TYPE "ST_PressDemoStationCfg"
VERSION : 0.1
   STRUCT
      "SchemaVersion" : UInt := 1;
      "RequireTwoHandStart" : Bool := TRUE;
      "TransferSettleTime" : Time := T#200ms;
      "PressSettleTime" : Time := T#300ms;
   END_STRUCT;
END_TYPE
